Fanuc KAREL source: ka00195.KL

-- PROVISIONAL review KL for V1013-1; original PC SHA256 3b054adbc48aadd97cbcc236d11275f41a3e9f713abdb223161383c1627ab8df
-- Incomplete behavior may be omitted. Consult companion uncertainty JSON. Do not deploy.
PROGRAM KA00195
%NOLOCKGROUP
-- UNRESOLVED_DECL SRC type=002017
-- UNRESOLVED_DECL DST type=002017
BEGIN
  -- UNRESOLVED_PC offsets 5-19; opcodes 22,22,1E
  -- UNRESOLVED_PC offsets 24-28; opcodes 7F
END KA00195
